FUNCTION F_Copy : BOOL
VAR_INPUT
    pSrc : POINTER TO DINT;
    pDst : POINTER TO DINT;
END_VAR

IF pSrc <> 0 THEN
    pDst^ := pSrc^; // PLCA-P005
END_IF

END_FUNCTION

(* stored: Version 1.1.0.1, ProductVersion 3.1.4024.12
   POU F_Copy: Id {00000000-0000-0000-0000-000000000001}, SpecialFunc None *)
